FUNCTION FC 1 : VOID
BEGIN
NETWORK
      L C#1000
END_FUNCTION
